Fanuc KAREL source: KX00014.KL

PROGRAM KX00014
%NOLOCKGROUP
VAR
  I: INTEGER
  J: INTEGER
  B: BOOLEAN
  F: FILE
  S: STRING[80]
  P: XYZWPR
BEGIN
  PURGE CONDITION[1]
END KX00014
